(* IEC 61131-3 sources: llm-plc-st-eval/data/definitivo/gemini-3.1-pro-preview/B3/zero_shot, 3 files *)

(* ---- ejec_1.st ---- *)
```iecst
FUNCTION_BLOCK FB_Contador
VAR_INPUT
    sensorPieza : BOOL; // Sensor fotoeléctrico (TRUE al detectar pieza)
    btnReset    : BOOL; // Botón para reiniciar la cuenta a cero
END_VAR

VAR_OUTPUT
    loteListo   : BOOL; // Se activa al llegar a 12 piezas
    cuenta      : INT;  // Número de piezas contadas
END_VAR

VAR
    flancoSensor : R_TRIG; // Detector de flanco de subida estándar IEC
END_VAR

// Detección del flanco de subida (transición de FALSE a TRUE) del sensor
flancoSensor(CLK := sensorPieza);

// Lógica de reinicio y conteo
IF btnReset THEN
    cuenta := 0; // Reinicia el contador
ELSIF flancoSensor.Q THEN
    cuenta := cuenta + 1; // Incrementa la cuenta por cada nueva pieza
END_IF;

// Evaluación del estado del lote (se desactiva automáticamente si cuenta < 12)
loteListo := (cuenta >= 12);

END_FUNCTION_BLOCK
```

(* ---- ejec_2.st ---- *)
```iecst
FUNCTION_BLOCK FB_Contador
VAR_INPUT
    sensorPieza : BOOL; // Sensor fotoeléctrico (TRUE al detectar pieza)
    btnReset    : BOOL; // Botón para reiniciar el contador
END_VAR

VAR_OUTPUT
    loteListo   : BOOL; // Se activa al llegar a 12 piezas
    cuenta      : INT;  // Número de piezas contadas
END_VAR

VAR
    flancoSensor : R_TRIG; // Bloque estándar para detectar flanco de subida
END_VAR

// Detectar transición de FALSE a TRUE en el sensor
flancoSensor(CLK := sensorPieza);

// Lógica de reinicio y conteo
IF btnReset THEN
    cuenta := 0; // Reiniciar cuenta
ELSIF flancoSensor.Q THEN
    cuenta := cuenta + 1; // Incrementar cuenta con cada nueva pieza
END_IF;

// Evaluar si el lote está completo (12 piezas)
// Al reiniciar la cuenta a 0, esta condición automáticamente desactiva loteListo
loteListo := (cuenta >= 12);

END_FUNCTION_BLOCK
```

(* ---- ejec_3.st ---- *)
```iecst
FUNCTION_BLOCK FB_Contador

VAR_INPUT
    sensorPieza : BOOL; // Entrada del sensor fotoeléctrico
    btnReset : BOOL;    // Botón para reiniciar el conteo y el lote
END_VAR

VAR_OUTPUT
    loteListo : BOOL;   // Se activa al llegar a 12 piezas
    cuenta : INT;       // Cantidad actual de piezas contadas
END_VAR

VAR
    flancoSensor : R_TRIG; // Instancia para detectar el flanco de subida
END_VAR

// Evaluar la transición de FALSE a TRUE del sensor
flancoSensor(CLK := sensorPieza);

// Lógica de reinicio y conteo
IF btnReset THEN
    cuenta := 0;
    loteListo := FALSE;
ELSIF flancoSensor.Q THEN
    cuenta := cuenta + 1;
END_IF;

// Lógica para activar la salida de lote completo
IF cuenta >= 12 THEN
    loteListo := TRUE;
END_IF;

END_FUNCTION_BLOCK
```
